Fanuc KAREL source: kd00053.compact.KL

PROGRAM KD00053
%STACKSIZE=65535
%PRIORITY=65535
%NOLOCKGROUP
VAR
I : INTEGER
J : INTEGER
B : BOOLEAN
R : REAL
S : STRING[80]
BEGIN
I=(J + 1)
END KD00053
